FUNCTION_BLOCK UCT_PreTratamento (* UCT Fast de tratamento preliminar + bomba de gordura - HidrycoLib *)
  (* Standard: 61499-2 *)
  (* Version 1.8, 12/11/2026, Hidryco, Hidryco, 1.8: termica da BombaGordura de volta a NF (cfgTermicaNF = TRUE: FALSE no campo = atuada), a pedido do usuario depois de corrigir os nomes dos symlinks (Pre_Tratamento1/2). 1.7: termica da BombaGordura invertida a pedido do usuario (cfgTermicaNF = FALSE: TRUE no campo = atuada). 1.6: IThis.STS_LIGADO, STS_AUTOMATICO (IO List da Nereda). 1.5: eventos da peneira rotativa na logica certa (liga manual em REQ_PEN_LIGA, velocidade em REQ_PEN_VEL, intermitente em REQ_PEN_INT). 1.4: simbolo sGordura (tanque de gordura e valvula de lavagem) para a tela do pre-tratamento. 1.3: sSkid reorganizado (tubos atras, equipamentos alinhados as portas), SymbolSize nos simbolos. 1.2: simbolo sSkid (desenho ISA-101 do skid, com os simbolos dos equipamentos e da bomba de gordura). 1.0: UCT Fast (tratamento preliminar, memorial PR-809) por Modbus TCP. Leitura pela configuracao de hardware (MODBUSGENTCPS + MODBUSRREG8/2 em 40005, 40013, 40081, 40101, 40116, 40127, 40136, 40151, 40161, 40230, 40500, 40508, 40516) nos symlinks ${PATH}mbW005..mbH517 (INT) e connStatusInt em ${PATH}mbConexao; escrita por MODBUSWREG1 em requestwrite nos symlinks ${PATH}mbEscW005..mbEscW017 e ${PATH}mbEscV101..mbEscV161 (INT), so quando o operador comanda. Equipamentos (sub-CATs UCT_Equipamento): Peneira, Bomba1, Bomba2, Valvula1, Valvula2, Compressor, Raspador, Rosca1, Rosca2. Disponibilidade pelo AND editavel (AND_UCT_OK e AND_DISPONIVEL); cadeia antHabilitada/antDisponivel -> stsBloqueioEEE. Bomba de gordura 200-BR-0x (Motor_Generico BombaGordura: E/S por ${PATH}BombaGordura.stsLocal/... e ATV: ComStatus direto em ${PATH}BombaGordura.stsFalhaComunicacao, o motor inverte) e valvula de lavagem ${PATH}cmdValvulaLavagem (BOOL). *)
  PACKAGE Hidryco.HidrycoLib;
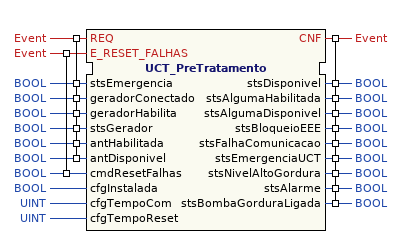
  EVENT_INPUT
    REQ WITH stsEmergencia, geradorConectado, geradorHabilita, stsGerador, antHabilitada, antDisponivel; (* Atualizacao do processo *)
    E_RESET_FALHAS WITH cmdResetFalhas; (* Reset pelo processo (UCT e bomba de gordura) com cmdResetFalhas = TRUE *)
  END_EVENT
  EVENT_OUTPUT
    CNF WITH stsDisponivel, stsAlgumaHabilitada, stsAlgumaDisponivel, stsBloqueioEEE, stsFalhaComunicacao, stsEmergenciaUCT, stsNivelAltoGordura, stsAlarme, stsBombaGorduraLigada; (* Disponibilidade, cadeia das UCTs e estados (so na mudanca) *)
  END_EVENT
  VAR_INPUT
    stsEmergencia : BOOL; (* Emergencia pelo processo: retira o comando da bomba de gordura e fecha a valvula de lavagem *)
    geradorConectado : BOOL := TRUE; (* A bomba de gordura pode ser alimentada pelo gerador *)
    geradorHabilita : BOOL; (* Bomba de gordura liberada para operar com a planta no gerador (HAB_UCT_200_0x do CAT Subestacao) *)
    stsGerador : BOOL; (* Planta alimentada pelo gerador *)
    antHabilitada : BOOL; (* Cadeia: alguma UCT anterior habilitada (stsAlgumaHabilitada da UCT anterior) *)
    antDisponivel : BOOL; (* Cadeia: alguma UCT anterior disponivel (stsAlgumaDisponivel da UCT anterior) *)
    cmdResetFalhas : BOOL; (* TRUE = reset (com o evento E_RESET_FALHAS) *)
    cfgInstalada : BOOL := TRUE; (* FALSE = UCT ainda nao existe em campo (sem comunicacao, sem alarmes, fora do bloqueio da EEE) *)
    cfgTempoCom : UINT := 10; (* Tempo (s) sem comunicacao com a UCT para confirmar a falha *)
    cfgTempoReset : UINT := 2; (* Tempo (s) do pulso de reset escrito na UCT (40005.3) *)
  END_VAR
  VAR_OUTPUT
    stsDisponivel : BOOL; (* UCT disponivel (saida do AND) *)
    stsAlgumaHabilitada : BOOL; (* Esta UCT ou alguma anterior habilitada *)
    stsAlgumaDisponivel : BOOL; (* Esta UCT ou alguma anterior disponivel *)
    stsBloqueioEEE : BOOL; (* Bloqueio do automatico da EEE Bruto: ha UCT habilitada e nenhuma disponivel *)
    stsFalhaComunicacao : BOOL; (* Falha de comunicacao com a UCT *)
    stsEmergenciaUCT : BOOL; (* Emergencia acionada na UCT *)
    stsNivelAltoGordura : BOOL; (* Nivel alto do tanque de gordura (UCT) *)
    stsAlarme : BOOL; (* Algum alarme da UCT *)
    stsBombaGorduraLigada : BOOL; (* Bomba de gordura ligada *)
  END_VAR
  FBS
    IThis : UCT_PreTratamento_HMI(QI := TRUE);
    plcStart1 : plcStart(Prio := 10);
    Logica : basicUCT;
    Tick : E_CYCLE(DT := T#1s);
    Leitura1 : SYMLINKMULTIVARDST_115C998103CD7017B(NAME1 := '$${PATH}mbW005', NAME2 := '$${PATH}mbW006', NAME3 := '$${PATH}mbW007', NAME4 := '$${PATH}mbW008', NAME5 := '$${PATH}mbW009', NAME6 := '$${PATH}mbW010', NAME7 := '$${PATH}mbW011', NAME8 := '$${PATH}mbW012', NAME9 := '$${PATH}mbW013', NAME10 := '$${PATH}mbW014', NAME11 := '$${PATH}mbW015', NAME12 := '$${PATH}mbW016', NAME13 := '$${PATH}mbW017', NAME14 := '$${PATH}mbW081', NAME15 := '$${PATH}mbW082', QI := TRUE); {SET_ATTRIBUTE(Configuration.GenericFBType.InterfaceParams, Runtime.System#I:=15;VALUE${I$}:INT,INT,INT,INT,INT,INT,INT,INT,INT,INT,INT,INT,INT,INT,INT)}
    Leitura2 : SYMLINKMULTIVARDST_115C998103CD7017B(NAME1 := '$${PATH}mbS101', NAME2 := '$${PATH}mbS106', NAME3 := '$${PATH}mbS116', NAME4 := '$${PATH}mbS117', NAME5 := '$${PATH}mbS121', NAME6 := '$${PATH}mbS122', NAME7 := '$${PATH}mbS127', NAME8 := '$${PATH}mbS132', NAME9 := '$${PATH}mbS136', NAME10 := '$${PATH}mbS137', NAME11 := '$${PATH}mbS141', NAME12 := '$${PATH}mbS142', NAME13 := '$${PATH}mbS151', NAME14 := '$${PATH}mbS152', NAME15 := '$${PATH}mbS161', QI := TRUE); {SET_ATTRIBUTE(Configuration.GenericFBType.InterfaceParams, Runtime.System#I:=15;VALUE${I$}:INT,INT,INT,INT,INT,INT,INT,INT,INT,INT,INT,INT,INT,INT,INT)}
    Leitura3 : SYMLINKMULTIVARDST_115C998103CD7017B(NAME1 := '$${PATH}mbS162', NAME2 := '$${PATH}mbW230', NAME3 := '$${PATH}mbH500', NAME4 := '$${PATH}mbH501', NAME5 := '$${PATH}mbH502', NAME6 := '$${PATH}mbH503', NAME7 := '$${PATH}mbH504', NAME8 := '$${PATH}mbH505', NAME9 := '$${PATH}mbH506', NAME10 := '$${PATH}mbH507', NAME11 := '$${PATH}mbH508', NAME12 := '$${PATH}mbH509', NAME13 := '$${PATH}mbH510', NAME14 := '$${PATH}mbH511', NAME15 := '$${PATH}mbH512', QI := TRUE); {SET_ATTRIBUTE(Configuration.GenericFBType.InterfaceParams, Runtime.System#I:=15;VALUE${I$}:INT,INT,INT,INT,INT,INT,INT,INT,INT,INT,INT,INT,INT,INT,INT)}
    Leitura4 : SYMLINKMULTIVARDST_15292F208F22048C1(NAME1 := '$${PATH}mbH513', NAME2 := '$${PATH}mbH514', NAME3 := '$${PATH}mbH515', NAME4 := '$${PATH}mbH516', QI := TRUE); {SET_ATTRIBUTE(Configuration.GenericFBType.InterfaceParams, Runtime.System#I:=4;VALUE${I$}:INT,INT,INT,INT)}
    Leitura5 : SYMLINKMULTIVARDST_5A03F112CD5D470(NAME1 := '$${PATH}mbH517', QI := TRUE); {SET_ATTRIBUTE(Configuration.GenericFBType.InterfaceParams, Runtime.System#I:=1;VALUE${I$}:INT)}
    Comunicacao : SYMLINKMULTIVARDST_5A03F112CD5D470(NAME1 := '$${PATH}mbConexao', QI := TRUE); {SET_ATTRIBUTE(Configuration.GenericFBType.InterfaceParams, Runtime.System#I:=1;VALUE${I$}:INT)}
    EscreveW005 : SYMLINKMULTIVARSRC_5A03F112CD5D470(NAME1 := '$${PATH}mbEscW005', QI := TRUE); {SET_ATTRIBUTE(Configuration.GenericFBType.InterfaceParams, Runtime.System#I:=1;VALUE${I$}:INT)}
    EscreveW006 : SYMLINKMULTIVARSRC_5A03F112CD5D470(NAME1 := '$${PATH}mbEscW006', QI := TRUE); {SET_ATTRIBUTE(Configuration.GenericFBType.InterfaceParams, Runtime.System#I:=1;VALUE${I$}:INT)}
    EscreveW007 : SYMLINKMULTIVARSRC_5A03F112CD5D470(NAME1 := '$${PATH}mbEscW007', QI := TRUE); {SET_ATTRIBUTE(Configuration.GenericFBType.InterfaceParams, Runtime.System#I:=1;VALUE${I$}:INT)}
    EscreveW008 : SYMLINKMULTIVARSRC_5A03F112CD5D470(NAME1 := '$${PATH}mbEscW008', QI := TRUE); {SET_ATTRIBUTE(Configuration.GenericFBType.InterfaceParams, Runtime.System#I:=1;VALUE${I$}:INT)}
    EscreveW009 : SYMLINKMULTIVARSRC_5A03F112CD5D470(NAME1 := '$${PATH}mbEscW009', QI := TRUE); {SET_ATTRIBUTE(Configuration.GenericFBType.InterfaceParams, Runtime.System#I:=1;VALUE${I$}:INT)}
    EscreveW010 : SYMLINKMULTIVARSRC_5A03F112CD5D470(NAME1 := '$${PATH}mbEscW010', QI := TRUE); {SET_ATTRIBUTE(Configuration.GenericFBType.InterfaceParams, Runtime.System#I:=1;VALUE${I$}:INT)}
    EscreveW011 : SYMLINKMULTIVARSRC_5A03F112CD5D470(NAME1 := '$${PATH}mbEscW011', QI := TRUE); {SET_ATTRIBUTE(Configuration.GenericFBType.InterfaceParams, Runtime.System#I:=1;VALUE${I$}:INT)}
    EscreveW012 : SYMLINKMULTIVARSRC_5A03F112CD5D470(NAME1 := '$${PATH}mbEscW012', QI := TRUE); {SET_ATTRIBUTE(Configuration.GenericFBType.InterfaceParams, Runtime.System#I:=1;VALUE${I$}:INT)}
    EscreveW013 : SYMLINKMULTIVARSRC_5A03F112CD5D470(NAME1 := '$${PATH}mbEscW013', QI := TRUE); {SET_ATTRIBUTE(Configuration.GenericFBType.InterfaceParams, Runtime.System#I:=1;VALUE${I$}:INT)}
    EscreveW014 : SYMLINKMULTIVARSRC_5A03F112CD5D470(NAME1 := '$${PATH}mbEscW014', QI := TRUE); {SET_ATTRIBUTE(Configuration.GenericFBType.InterfaceParams, Runtime.System#I:=1;VALUE${I$}:INT)}
    EscreveW015 : SYMLINKMULTIVARSRC_5A03F112CD5D470(NAME1 := '$${PATH}mbEscW015', QI := TRUE); {SET_ATTRIBUTE(Configuration.GenericFBType.InterfaceParams, Runtime.System#I:=1;VALUE${I$}:INT)}
    EscreveW016 : SYMLINKMULTIVARSRC_5A03F112CD5D470(NAME1 := '$${PATH}mbEscW016', QI := TRUE); {SET_ATTRIBUTE(Configuration.GenericFBType.InterfaceParams, Runtime.System#I:=1;VALUE${I$}:INT)}
    EscreveW017 : SYMLINKMULTIVARSRC_5A03F112CD5D470(NAME1 := '$${PATH}mbEscW017', QI := TRUE); {SET_ATTRIBUTE(Configuration.GenericFBType.InterfaceParams, Runtime.System#I:=1;VALUE${I$}:INT)}
    EscreveV101 : SYMLINKMULTIVARSRC_5A03F112CD5D470(NAME1 := '$${PATH}mbEscV101', QI := TRUE); {SET_ATTRIBUTE(Configuration.GenericFBType.InterfaceParams, Runtime.System#I:=1;VALUE${I$}:INT)}
    EscreveV116 : SYMLINKMULTIVARSRC_5A03F112CD5D470(NAME1 := '$${PATH}mbEscV116', QI := TRUE); {SET_ATTRIBUTE(Configuration.GenericFBType.InterfaceParams, Runtime.System#I:=1;VALUE${I$}:INT)}
    EscreveV121 : SYMLINKMULTIVARSRC_5A03F112CD5D470(NAME1 := '$${PATH}mbEscV121', QI := TRUE); {SET_ATTRIBUTE(Configuration.GenericFBType.InterfaceParams, Runtime.System#I:=1;VALUE${I$}:INT)}
    EscreveV136 : SYMLINKMULTIVARSRC_5A03F112CD5D470(NAME1 := '$${PATH}mbEscV136', QI := TRUE); {SET_ATTRIBUTE(Configuration.GenericFBType.InterfaceParams, Runtime.System#I:=1;VALUE${I$}:INT)}
    EscreveV141 : SYMLINKMULTIVARSRC_5A03F112CD5D470(NAME1 := '$${PATH}mbEscV141', QI := TRUE); {SET_ATTRIBUTE(Configuration.GenericFBType.InterfaceParams, Runtime.System#I:=1;VALUE${I$}:INT)}
    EscreveV151 : SYMLINKMULTIVARSRC_5A03F112CD5D470(NAME1 := '$${PATH}mbEscV151', QI := TRUE); {SET_ATTRIBUTE(Configuration.GenericFBType.InterfaceParams, Runtime.System#I:=1;VALUE${I$}:INT)}
    EscreveV161 : SYMLINKMULTIVARSRC_5A03F112CD5D470(NAME1 := '$${PATH}mbEscV161', QI := TRUE); {SET_ATTRIBUTE(Configuration.GenericFBType.InterfaceParams, Runtime.System#I:=1;VALUE${I$}:INT)}
    ValvulaLavagem : SYMLINKMULTIVARSRC_1559B0FF8170C9BA0(NAME1 := '$${PATH}cmdValvulaLavagem', QI := TRUE); {SET_ATTRIBUTE(Configuration.GenericFBType.InterfaceParams, Runtime.System#I:=1;VALUE${I$}:BOOL)}
    AND_UCT_OK : AND_1122770BAB85676D3; {SET_ATTRIBUTE(Configuration.GenericFBType.InterfaceParams, Runtime.Standard#CNT:=3)}
    AND_DISPONIVEL : AND_1122770BAB85676D3; {SET_ATTRIBUTE(Configuration.GenericFBType.InterfaceParams, Runtime.Standard#CNT:=3)}
    Bomba_Higienizacao1 : UCT_Equipamento(pin_6729E072E11CC02E := TRUE, pin_B3CA2188BE2BF3D0 := FALSE, pin_E5B528FA2A3E5A83 := FALSE);
    Bomba_Higienizacao2 : UCT_Equipamento(pin_6729E072E11CC02E := TRUE, pin_B3CA2188BE2BF3D0 := FALSE, pin_E5B528FA2A3E5A83 := FALSE);
    Valvula_Higienizacao1 : UCT_Equipamento(pin_6729E072E11CC02E := FALSE, pin_B3CA2188BE2BF3D0 := FALSE, pin_E5B528FA2A3E5A83 := FALSE);
    Valvula_Higienizacao2 : UCT_Equipamento(pin_6729E072E11CC02E := FALSE, pin_B3CA2188BE2BF3D0 := FALSE, pin_E5B528FA2A3E5A83 := FALSE);
    Compressor1 : UCT_Equipamento(pin_6729E072E11CC02E := TRUE, pin_B3CA2188BE2BF3D0 := FALSE, pin_E5B528FA2A3E5A83 := FALSE);
    Raspador_Gordura1 : UCT_Equipamento(pin_6729E072E11CC02E := TRUE, pin_B3CA2188BE2BF3D0 := TRUE, pin_E5B528FA2A3E5A83 := TRUE);
    Rosca1Horizontal : UCT_Equipamento(pin_6729E072E11CC02E := TRUE, pin_B3CA2188BE2BF3D0 := TRUE, pin_E5B528FA2A3E5A83 := TRUE);
    Rosca2Inclinada : UCT_Equipamento(pin_6729E072E11CC02E := TRUE, pin_B3CA2188BE2BF3D0 := TRUE, pin_E5B528FA2A3E5A83 := TRUE);
    BombaGordura : Motor_Generico(pin_63EFEFB7C85EC93E := TRUE, pin_66763E13F70A4420 := TRUE, pin_D34C88BE7FFF3208 := TRUE, pin_39489193B7758574 := 600.0);
    AlarmeCom : ALARM_BIT(TYPE := 1, ACKTYPE_1 := 2, ACTIVE := TRUE); {SET_ATTRIBUTE(HMI.AlarmText, UCT sem comunicação)}
    AlarmeEmergencia : ALARM_BIT(TYPE := 1, ACKTYPE_1 := 2, ACTIVE := TRUE); {SET_ATTRIBUTE(HMI.AlarmText, Emergência acionada na UCT)}
    AlarmeDefPEN : ALARM_BIT(TYPE := 1, ACKTYPE_1 := 2, ACTIVE := TRUE); {SET_ATTRIBUTE(HMI.AlarmText, Defeito na peneira rotativa)}
    AlarmeDefB1 : ALARM_BIT(TYPE := 1, ACKTYPE_1 := 2, ACTIVE := TRUE); {SET_ATTRIBUTE(HMI.AlarmText, Defeito na bomba 1 de higienização da peneira)}
    AlarmeDefB2 : ALARM_BIT(TYPE := 1, ACKTYPE_1 := 2, ACTIVE := TRUE); {SET_ATTRIBUTE(HMI.AlarmText, Defeito na bomba 2 de higienização da peneira)}
    AlarmeDefCMP : ALARM_BIT(TYPE := 1, ACKTYPE_1 := 2, ACTIVE := TRUE); {SET_ATTRIBUTE(HMI.AlarmText, Defeito no compressor de ar)}
    AlarmeDefRSP : ALARM_BIT(TYPE := 1, ACKTYPE_1 := 2, ACTIVE := TRUE); {SET_ATTRIBUTE(HMI.AlarmText, Defeito no raspador de gordura)}
    AlarmeDefR1 : ALARM_BIT(TYPE := 1, ACKTYPE_1 := 2, ACTIVE := TRUE); {SET_ATTRIBUTE(HMI.AlarmText, Defeito na rosca 1 (horizontal))}
    AlarmeDefR2 : ALARM_BIT(TYPE := 1, ACKTYPE_1 := 2, ACTIVE := TRUE); {SET_ATTRIBUTE(HMI.AlarmText, Defeito na rosca 2 (inclinada))}
    AlarmeNivelAgua : ALARM_BIT(TYPE := 1, ACKTYPE_1 := 2, ACTIVE := TRUE); {SET_ATTRIBUTE(HMI.AlarmText, Nível baixo no tanque de água de higienização)} {SET_ATTRIBUTE(HMI.AlarmClass, Warning)}
    AlarmeNivelPeneira : ALARM_BIT(TYPE := 1, ACKTYPE_1 := 2, ACTIVE := TRUE); {SET_ATTRIBUTE(HMI.AlarmText, Nível alto na peneira)} {SET_ATTRIBUTE(HMI.AlarmClass, Warning)}
    Peneira_Rotativa1 : UCT_Equipamento(pin_6729E072E11CC02E := TRUE, pin_B3CA2188BE2BF3D0 := TRUE, pin_E5B528FA2A3E5A83 := FALSE);
  END_FBS
  EVENT_CONNECTIONS
    plcStart1.FIRST_INIT TO IThis.7731B1FFA94C6332;
    plcStart1.REDO_INIT TO IThis.7731B1FFA94C6332;
    IThis.BE90C28BEC8DBAC0 TO Logica.3C5B6DD981EA9EF0;
    Logica.416B84A41F220B84 TO Tick.START;
    Logica.416B84A41F220B84 TO Leitura1.INIT;
    Logica.416B84A41F220B84 TO Leitura2.INIT;
    Logica.416B84A41F220B84 TO Leitura3.INIT;
    Logica.416B84A41F220B84 TO Leitura4.INIT;
    Logica.416B84A41F220B84 TO Leitura5.INIT;
    Logica.416B84A41F220B84 TO Comunicacao.INIT;
    Logica.416B84A41F220B84 TO EscreveW005.INIT;
    Logica.416B84A41F220B84 TO EscreveW006.INIT;
    Logica.416B84A41F220B84 TO EscreveW007.INIT;
    Logica.416B84A41F220B84 TO EscreveW008.INIT;
    Logica.416B84A41F220B84 TO EscreveW009.INIT;
    Logica.416B84A41F220B84 TO EscreveW010.INIT;
    Logica.416B84A41F220B84 TO EscreveW011.INIT;
    Logica.416B84A41F220B84 TO EscreveW012.INIT;
    Logica.416B84A41F220B84 TO EscreveW013.INIT;
    Logica.416B84A41F220B84 TO EscreveW014.INIT;
    Logica.416B84A41F220B84 TO EscreveW015.INIT;
    Logica.416B84A41F220B84 TO EscreveW016.INIT;
    Logica.416B84A41F220B84 TO EscreveW017.INIT;
    Logica.416B84A41F220B84 TO EscreveV101.INIT;
    Logica.416B84A41F220B84 TO EscreveV116.INIT;
    Logica.416B84A41F220B84 TO EscreveV121.INIT;
    Logica.416B84A41F220B84 TO EscreveV136.INIT;
    Logica.416B84A41F220B84 TO EscreveV141.INIT;
    Logica.416B84A41F220B84 TO EscreveV151.INIT;
    Logica.416B84A41F220B84 TO EscreveV161.INIT;
    Logica.416B84A41F220B84 TO ValvulaLavagem.INIT;
    Logica.416B84A41F220B84 TO AlarmeCom.INIT;
    AlarmeCom.INITO TO AlarmeCom.REQ_INITDATA;
    AlarmeCom.CNF_INITDATA TO AlarmeCom.ACTIVATE;
    AlarmeCom.INITO TO AlarmeEmergencia.INIT;
    AlarmeEmergencia.INITO TO AlarmeEmergencia.REQ_INITDATA;
    AlarmeEmergencia.CNF_INITDATA TO AlarmeEmergencia.ACTIVATE;
    AlarmeEmergencia.INITO TO AlarmeDefPEN.INIT;
    AlarmeDefPEN.INITO TO AlarmeDefPEN.REQ_INITDATA;
    AlarmeDefPEN.CNF_INITDATA TO AlarmeDefPEN.ACTIVATE;
    AlarmeDefPEN.INITO TO AlarmeDefB1.INIT;
    AlarmeDefB1.INITO TO AlarmeDefB1.REQ_INITDATA;
    AlarmeDefB1.CNF_INITDATA TO AlarmeDefB1.ACTIVATE;
    AlarmeDefB1.INITO TO AlarmeDefB2.INIT;
    AlarmeDefB2.INITO TO AlarmeDefB2.REQ_INITDATA;
    AlarmeDefB2.CNF_INITDATA TO AlarmeDefB2.ACTIVATE;
    AlarmeDefB2.INITO TO AlarmeDefCMP.INIT;
    AlarmeDefCMP.INITO TO AlarmeDefCMP.REQ_INITDATA;
    AlarmeDefCMP.CNF_INITDATA TO AlarmeDefCMP.ACTIVATE;
    AlarmeDefCMP.INITO TO AlarmeDefRSP.INIT;
    AlarmeDefRSP.INITO TO AlarmeDefRSP.REQ_INITDATA;
    AlarmeDefRSP.CNF_INITDATA TO AlarmeDefRSP.ACTIVATE;
    AlarmeDefRSP.INITO TO AlarmeDefR1.INIT;
    AlarmeDefR1.INITO TO AlarmeDefR1.REQ_INITDATA;
    AlarmeDefR1.CNF_INITDATA TO AlarmeDefR1.ACTIVATE;
    AlarmeDefR1.INITO TO AlarmeDefR2.INIT;
    AlarmeDefR2.INITO TO AlarmeDefR2.REQ_INITDATA;
    AlarmeDefR2.CNF_INITDATA TO AlarmeDefR2.ACTIVATE;
    AlarmeDefR2.INITO TO AlarmeNivelAgua.INIT;
    AlarmeNivelAgua.INITO TO AlarmeNivelAgua.REQ_INITDATA;
    AlarmeNivelAgua.CNF_INITDATA TO AlarmeNivelAgua.ACTIVATE;
    AlarmeNivelAgua.INITO TO AlarmeNivelPeneira.INIT;
    AlarmeNivelPeneira.INITO TO AlarmeNivelPeneira.REQ_INITDATA;
    AlarmeNivelPeneira.CNF_INITDATA TO AlarmeNivelPeneira.ACTIVATE;
    AlarmeNivelPeneira.INITO TO plcStart1.ACK_FIRST;
    AlarmeNivelPeneira.INITO TO IThis.BF3BAA6EB0D69F6F;
    Leitura1.CNF TO Logica.86B21E575F925410;
    Leitura2.CNF TO Logica.ACF117E29FC3AC1C;
    Leitura3.CNF TO Logica.FD034B0BBE440D40;
    Leitura4.CNF TO Logica.729388FCDFDF68AE;
    Leitura5.CNF TO Logica.96AC3F0A2629C81D;
    Comunicacao.CNF TO Logica.4327DB3EB2D5D05C;
    Logica.11F41745985917DF TO EscreveW005.REQ;
    Logica.E9DD31896C582136 TO EscreveW006.REQ;
    Logica.E928AC62D8378E2E TO EscreveW007.REQ;
    Logica.8C6CC9C5F833000C TO EscreveW008.REQ;
    Logica.10A819F294BECD61 TO EscreveW009.REQ;
    Logica.CCE6CEE36384A6FD TO EscreveW010.REQ;
    Logica.48F5F46EFA41CB2E TO EscreveW011.REQ;
    Logica.FB2D821A4BBF6B61 TO EscreveW012.REQ;
    Logica.6F9E0D27072C9DCA TO EscreveW013.REQ;
    Logica.3830C851999B1CA8 TO EscreveW014.REQ;
    Logica.91DFFB362B8ECB72 TO EscreveW015.REQ;
    Logica.D8E5B77061056FA5 TO EscreveW016.REQ;
    Logica.67B496F21A680217 TO EscreveW017.REQ;
    Logica.2DC67FC3F907B62C TO EscreveV101.REQ;
    Logica.9697531BFDFDAA11 TO EscreveV116.REQ;
    Logica.EA10A30027EF1458 TO EscreveV121.REQ;
    Logica.76B63473D5644862 TO EscreveV136.REQ;
    Logica.E8A88BE3B83ED632 TO EscreveV141.REQ;
    Logica.FCC1975F18BB837D TO EscreveV151.REQ;
    Logica.D44CECCDCDAFDF05 TO EscreveV161.REQ;
    Logica.8621D711C765D74F TO ValvulaLavagem.REQ;
    Logica.A0C13DD0452107CB TO Bomba_Higienizacao1.70A516C5CA4155CA;
    Bomba_Higienizacao1.0ECDAB45E7B0C5AF TO Logica.9D9E81ADADCAA296;
    Bomba_Higienizacao1.2D7A148B2A7AA879 TO Logica.E34661574BF84379;
    Logica.A0C13DD0452107CB TO Bomba_Higienizacao2.70A516C5CA4155CA;
    Bomba_Higienizacao2.0ECDAB45E7B0C5AF TO Logica.D87E7B2D8E293BB6;
    Bomba_Higienizacao2.2D7A148B2A7AA879 TO Logica.7CA1C2A34CD31341;
    Logica.A0C13DD0452107CB TO Valvula_Higienizacao1.70A516C5CA4155CA;
    Valvula_Higienizacao1.0ECDAB45E7B0C5AF TO Logica.CF56824B76A4E51B;
    Logica.A0C13DD0452107CB TO Valvula_Higienizacao2.70A516C5CA4155CA;
    Valvula_Higienizacao2.0ECDAB45E7B0C5AF TO Logica.F75EA032D1A6B02C;
    Logica.A0C13DD0452107CB TO Compressor1.70A516C5CA4155CA;
    Compressor1.0ECDAB45E7B0C5AF TO Logica.548C5ECAC6439F23;
    Compressor1.2D7A148B2A7AA879 TO Logica.D33EB6DFF7EADA48;
    Logica.A0C13DD0452107CB TO Raspador_Gordura1.70A516C5CA4155CA;
    Raspador_Gordura1.0ECDAB45E7B0C5AF TO Logica.4F24C39CA1B377DA;
    Raspador_Gordura1.453EBF0958E76CD5 TO Logica.25A416A6D88DD0BD;
    Raspador_Gordura1.D9A88CBEE21DBA8E TO Logica.2DDC9EB582C567B6;
    Raspador_Gordura1.2D7A148B2A7AA879 TO Logica.E445565C572BE9AB;
    Logica.A0C13DD0452107CB TO Rosca1Horizontal.70A516C5CA4155CA;
    Rosca1Horizontal.0ECDAB45E7B0C5AF TO Logica.B6026660A2849366;
    Rosca1Horizontal.453EBF0958E76CD5 TO Logica.38389BFD6E07A057;
    Rosca1Horizontal.D9A88CBEE21DBA8E TO Logica.460B0CE006F8F781;
    Rosca1Horizontal.2D7A148B2A7AA879 TO Logica.9798AA2801C41B49;
    Logica.A0C13DD0452107CB TO Rosca2Inclinada.70A516C5CA4155CA;
    Rosca2Inclinada.0ECDAB45E7B0C5AF TO Logica.05FCFC0A4F34DAC5;
    Rosca2Inclinada.453EBF0958E76CD5 TO Logica.917F967EEA65C256;
    Rosca2Inclinada.D9A88CBEE21DBA8E TO Logica.F6429B88CEB00ADB;
    Rosca2Inclinada.2D7A148B2A7AA879 TO Logica.66FC9636E69253EA;
    IThis.1F1F8302525DDF94 TO Logica.60A9FA7D1B9019D9;
    IThis.1EA45A01E944042C TO Logica.10C669586AF9B729;
    IThis.6BDBFED6495F25F4 TO Logica.70D47E2D73B66C31;
    IThis.734C7A77C68CFD95 TO Logica.10434994C0931297;
    IThis.E2F5EBA7E91047EB TO Logica.4287AE5C00B681B1;
    IThis.CA131EB7F5B48041 TO Logica.8858219971D3BAD6;
    IThis.09F2CE520A7CB40A TO Logica.B055BD39F7E10E53;
    IThis.74FD7728297A1739 TO Logica.8B3CC5BA21742708;
    IThis.36C4ED263F60138F TO Logica.01DDB779929E0BD3;
    IThis.313AA7AFD2DEA98C TO Logica.FF42D335F0EB104F;
    E_RESET_FALHAS TO Logica.F6EC819575FB3804;
    REQ TO Logica.75410FBD6637F3BE;
    REQ TO BombaGordura.21070E4B73BFECDC;
    Tick.EO TO Logica.41222487C8D9CF7D;
    Logica.A4E8AA815C7798D0 TO CNF;
    Logica.B1173782F7B0D885 TO IThis.4D2C1FBBFC38ACE6;
    Logica.4C6FF34A6B3F84FA TO AND_UCT_OK.REQ;
    AND_UCT_OK.CNF TO AND_DISPONIVEL.REQ;
    AND_DISPONIVEL.CNF TO Logica.B4B1263914B085C1;
    Logica.31FE10FED34E3AE0 TO BombaGordura.21070E4B73BFECDC;
    BombaGordura.9D4F26EE27EDF5B9 TO Logica.7F4121B3EAF345EF;
    BombaGordura.9D4F26EE27EDF5B9 TO CNF;
    Logica.61B5851DEAB87FC2 TO BombaGordura.BA30A65ADDA4ECC3;
    Logica.B2C6B3F912408F66 TO AlarmeCom.REQ;
    Logica.B2C6B3F912408F66 TO AlarmeEmergencia.REQ;
    Logica.B2C6B3F912408F66 TO AlarmeDefPEN.REQ;
    Logica.B2C6B3F912408F66 TO AlarmeDefB1.REQ;
    Logica.B2C6B3F912408F66 TO AlarmeDefB2.REQ;
    Logica.B2C6B3F912408F66 TO AlarmeDefCMP.REQ;
    Logica.B2C6B3F912408F66 TO AlarmeDefRSP.REQ;
    Logica.B2C6B3F912408F66 TO AlarmeDefR1.REQ;
    Logica.B2C6B3F912408F66 TO AlarmeDefR2.REQ;
    Logica.B2C6B3F912408F66 TO AlarmeNivelAgua.REQ;
    Logica.B2C6B3F912408F66 TO AlarmeNivelPeneira.REQ;
    AlarmeCom.IND_1 TO IThis.4D2C1FBBFC38ACE6;
    AlarmeEmergencia.IND_1 TO IThis.4D2C1FBBFC38ACE6;
    AlarmeDefPEN.IND_1 TO IThis.4D2C1FBBFC38ACE6;
    AlarmeDefB1.IND_1 TO IThis.4D2C1FBBFC38ACE6;
    AlarmeDefB2.IND_1 TO IThis.4D2C1FBBFC38ACE6;
    AlarmeDefCMP.IND_1 TO IThis.4D2C1FBBFC38ACE6;
    AlarmeDefRSP.IND_1 TO IThis.4D2C1FBBFC38ACE6;
    AlarmeDefR1.IND_1 TO IThis.4D2C1FBBFC38ACE6;
    AlarmeDefR2.IND_1 TO IThis.4D2C1FBBFC38ACE6;
    AlarmeNivelAgua.IND_1 TO IThis.4D2C1FBBFC38ACE6;
    AlarmeNivelPeneira.IND_1 TO IThis.4D2C1FBBFC38ACE6;
    IThis.74FD7728297A1739 TO AlarmeCom.ACK_C1;
    IThis.74FD7728297A1739 TO AlarmeEmergencia.ACK_C1;
    IThis.74FD7728297A1739 TO AlarmeDefPEN.ACK_C1;
    IThis.74FD7728297A1739 TO AlarmeDefB1.ACK_C1;
    IThis.74FD7728297A1739 TO AlarmeDefB2.ACK_C1;
    IThis.74FD7728297A1739 TO AlarmeDefCMP.ACK_C1;
    IThis.74FD7728297A1739 TO AlarmeDefRSP.ACK_C1;
    IThis.74FD7728297A1739 TO AlarmeDefR1.ACK_C1;
    IThis.74FD7728297A1739 TO AlarmeDefR2.ACK_C1;
    IThis.74FD7728297A1739 TO AlarmeNivelAgua.ACK_C1;
    IThis.74FD7728297A1739 TO AlarmeNivelPeneira.ACK_C1;
    E_RESET_FALHAS TO AlarmeCom.ACK_C1;
    E_RESET_FALHAS TO AlarmeEmergencia.ACK_C1;
    E_RESET_FALHAS TO AlarmeDefPEN.ACK_C1;
    E_RESET_FALHAS TO AlarmeDefB1.ACK_C1;
    E_RESET_FALHAS TO AlarmeDefB2.ACK_C1;
    E_RESET_FALHAS TO AlarmeDefCMP.ACK_C1;
    E_RESET_FALHAS TO AlarmeDefRSP.ACK_C1;
    E_RESET_FALHAS TO AlarmeDefR1.ACK_C1;
    E_RESET_FALHAS TO AlarmeDefR2.ACK_C1;
    E_RESET_FALHAS TO AlarmeNivelAgua.ACK_C1;
    E_RESET_FALHAS TO AlarmeNivelPeneira.ACK_C1;
    Logica.A4E8AA815C7798D0 TO Peneira_Rotativa1.70A516C5CA4155CA;
    Logica.B1173782F7B0D885 TO Peneira_Rotativa1.70A516C5CA4155CA;
    Logica.A0C13DD0452107CB TO Peneira_Rotativa1.70A516C5CA4155CA;
    Logica.4C6FF34A6B3F84FA TO Peneira_Rotativa1.70A516C5CA4155CA;
    Logica.B2C6B3F912408F66 TO Peneira_Rotativa1.70A516C5CA4155CA;
    Logica.31FE10FED34E3AE0 TO Peneira_Rotativa1.70A516C5CA4155CA;
    Logica.8621D711C765D74F TO Peneira_Rotativa1.70A516C5CA4155CA;
    Logica.61B5851DEAB87FC2 TO Peneira_Rotativa1.70A516C5CA4155CA;
    Peneira_Rotativa1.0ECDAB45E7B0C5AF TO Logica.F5A0AE6E537529F5;
    Peneira_Rotativa1.2D7A148B2A7AA879 TO Logica.4A489282C873CE35;
    Peneira_Rotativa1.453EBF0958E76CD5 TO Logica.CB1FF06E5DD10F71;
  END_CONNECTIONS
  DATA_CONNECTIONS
    cfgInstalada TO Logica.B84AF20A00A0FEAB;
    cfgTempoCom TO Logica.2D0DECC616DD4E29;
    cfgTempoReset TO Logica.6F72EF7A9957D9B1;
    cmdResetFalhas TO Logica.F64D45B3992C3082;
    antHabilitada TO Logica.CF63D4AF765659C1;
    antDisponivel TO Logica.9756EA9EC3EE5693;
    stsEmergencia TO Logica.BCC8272ACE7AC349;
    Leitura1.VALUE1 TO Logica.2AF241D1E0537909;
    Leitura1.VALUE2 TO Logica.EB87F4844550BF0A;
    Leitura1.VALUE3 TO Logica.702CACE592B586EC;
    Leitura1.VALUE4 TO Logica.00E434C4D2FCE1E2;
    Leitura1.VALUE5 TO Logica.216DC8D1B0130B70;
    Leitura1.VALUE6 TO Logica.E92E8124C98345A8;
    Leitura1.VALUE7 TO Logica.5702FCE80FD9232F;
    Leitura1.VALUE8 TO Logica.2C198397DC93FDE4;
    Leitura1.VALUE9 TO Logica.8DC0D656670A81AF;
    Leitura1.VALUE10 TO Logica.FF2A6CB505BDEEED;
    Leitura1.VALUE11 TO Logica.29D39A9131350120;
    Leitura1.VALUE12 TO Logica.5047554D33D25508;
    Leitura1.VALUE13 TO Logica.6213901E687BF582;
    Leitura1.VALUE14 TO Logica.805F5AA59EEEC2D4;
    Leitura1.VALUE15 TO Logica.8AF7D7600739FBD8;
    Leitura2.VALUE1 TO Logica.CBA17D927032CBD4;
    Leitura2.VALUE2 TO Logica.E81009FF89B5BC15;
    Leitura2.VALUE3 TO Logica.FDB62ADC45542E9E;
    Leitura2.VALUE4 TO Logica.6D9544B2D05EE83A;
    Leitura2.VALUE5 TO Logica.EAC2F7A409142C5D;
    Leitura2.VALUE6 TO Logica.2873DE3B6BFE44C9;
    Leitura2.VALUE7 TO Logica.DB13AC717A8B7662;
    Leitura2.VALUE8 TO Logica.4D5D876EB3A7F171;
    Leitura2.VALUE9 TO Logica.51DA211617F1996B;
    Leitura2.VALUE10 TO Logica.97151C90B367E8DC;
    Leitura2.VALUE11 TO Logica.EEFE5F1EF8383B49;
    Leitura2.VALUE12 TO Logica.62F04539174C591F;
    Leitura2.VALUE13 TO Logica.02097632451711DE;
    Leitura2.VALUE14 TO Logica.7991843F9B2D5590;
    Leitura2.VALUE15 TO Logica.DDA25525CB8A7B4D;
    Leitura3.VALUE1 TO Logica.111326FFB7350BF0;
    Leitura3.VALUE2 TO Logica.605236348EF76178;
    Leitura3.VALUE3 TO Logica.009C88AD569306A2;
    Leitura3.VALUE4 TO Logica.A0B989F0831D5C46;
    Leitura3.VALUE5 TO Logica.C7387B9A6FCCB81F;
    Leitura3.VALUE6 TO Logica.E47649B3DC153190;
    Leitura3.VALUE7 TO Logica.3553691F126CE1B5;
    Leitura3.VALUE8 TO Logica.0A36A58BDBBC0471;
    Leitura3.VALUE9 TO Logica.42520E00029B280F;
    Leitura3.VALUE10 TO Logica.B3A245D474F32D30;
    Leitura3.VALUE11 TO Logica.FDF3C709AEBF1C84;
    Leitura3.VALUE12 TO Logica.25EE4A659CDB8B19;
    Leitura3.VALUE13 TO Logica.8E1D474EDFE3E373;
    Leitura3.VALUE14 TO Logica.A05F827665BFFF1E;
    Leitura3.VALUE15 TO Logica.DE0C347B4E1AA668;
    Leitura4.VALUE1 TO Logica.BE7F6B173ECEF46F;
    Leitura4.VALUE2 TO Logica.5FDC3C3D54E86285;
    Leitura4.VALUE3 TO Logica.D1FE5B095A8ACDE9;
    Leitura4.VALUE4 TO Logica.8A95E69557A2E9BE;
    Leitura5.VALUE1 TO Logica.ED8792C392F4F103;
    Comunicacao.VALUE1 TO Logica.8E65120B34D38BDE;
    Logica.48B51513B83DEAC1 TO EscreveW005.VALUE1;
    Logica.ABE25A7B6D246024 TO EscreveW006.VALUE1;
    Logica.332BB6C4B414C757 TO EscreveW007.VALUE1;
    Logica.5FF35C3FF4051574 TO EscreveW008.VALUE1;
    Logica.7BCA7ABE5B2A80CB TO EscreveW009.VALUE1;
    Logica.EE8A41D2485DFDB4 TO EscreveW010.VALUE1;
    Logica.A2EA9BE38D7D6BAA TO EscreveW011.VALUE1;
    Logica.126C934AB0F6DBFE TO EscreveW012.VALUE1;
    Logica.73DD8991441412AC TO EscreveW013.VALUE1;
    Logica.DE2C0333DCDCC77C TO EscreveW014.VALUE1;
    Logica.8B46394DF76CFFD8 TO EscreveW015.VALUE1;
    Logica.B5B936F289F2140E TO EscreveW016.VALUE1;
    Logica.96F874CA969849BC TO EscreveW017.VALUE1;
    Logica.93EC120EF49D8A9B TO EscreveV101.VALUE1;
    Logica.B84F5A34C7CB0F43 TO EscreveV116.VALUE1;
    Logica.2EEB0ECC5C70DFC8 TO EscreveV121.VALUE1;
    Logica.A95766D7DCAD36EA TO EscreveV136.VALUE1;
    Logica.D451279D5E50FC08 TO EscreveV141.VALUE1;
    Logica.D04BD37BABA3A53F TO EscreveV151.VALUE1;
    Logica.77B5D89A59E485CC TO EscreveV161.VALUE1;
    Logica.97A930D5B8996F70 TO ValvulaLavagem.VALUE1;
    Logica.4FE6015A2477CFC9 TO AND_UCT_OK.IN1;
    Logica.3836FD4FBDBFBB63 TO AND_UCT_OK.IN2;
    Logica.CFDFC80ABF4D39D0 TO AND_UCT_OK.IN3;
    AND_UCT_OK.OUT TO AND_DISPONIVEL.IN1;
    Logica.9719C72C2028949E TO AND_DISPONIVEL.IN2;
    Logica.EAECF18552174CCF TO AND_DISPONIVEL.IN3;
    AND_DISPONIVEL.OUT TO Logica.907F6462227B081B;
    Logica.9F5A0BAAA6BA36FB TO Bomba_Higienizacao1.93B31B867A532500;
    Logica.B0882E75048E56C8 TO Bomba_Higienizacao1.98FD5EAA90BD9629;
    Logica.F433D77752764E72 TO Bomba_Higienizacao1.96E48787F8AC58C3;
    Logica.BB50EA5A17772016 TO Bomba_Higienizacao1.CC220F735371196B;
    Logica.6D499885ADD13F89 TO Bomba_Higienizacao1.33285C93B9AAB2BC;
    Logica.6F1E502C9B6CF2B2 TO Bomba_Higienizacao1.3F39B194DE4581AB;
    Logica.B8856E3515E1335F TO Bomba_Higienizacao1.F6AE4997ED76CC8B;
    Logica.48FD745C0144715F TO Bomba_Higienizacao1.0E2695E0A2003068;
    Bomba_Higienizacao1.074D328E856330C0 TO Logica.C19AEC3805E7291E;
    Bomba_Higienizacao1.520AB5A4EADBD8AE TO Logica.878937D8CA59CE95;
    Logica.26DA29A2F44AB1D9 TO Bomba_Higienizacao2.93B31B867A532500;
    Logica.AE4A01B00246A9BC TO Bomba_Higienizacao2.98FD5EAA90BD9629;
    Logica.49B62932E0024FCB TO Bomba_Higienizacao2.96E48787F8AC58C3;
    Logica.C62B70166A0883C7 TO Bomba_Higienizacao2.CC220F735371196B;
    Logica.3229D99A95CB4D5D TO Bomba_Higienizacao2.33285C93B9AAB2BC;
    Logica.AC94358F5B25F765 TO Bomba_Higienizacao2.3F39B194DE4581AB;
    Logica.8F6F2CB2BBCF9FC3 TO Bomba_Higienizacao2.F6AE4997ED76CC8B;
    Logica.4FF14F19D4AA0DEA TO Bomba_Higienizacao2.0E2695E0A2003068;
    Bomba_Higienizacao2.074D328E856330C0 TO Logica.6F688A786E95C4D1;
    Bomba_Higienizacao2.520AB5A4EADBD8AE TO Logica.3A9274E19001885E;
    Logica.9594942602D571EA TO Valvula_Higienizacao1.93B31B867A532500;
    Logica.3A38DC7CA6958C9C TO Valvula_Higienizacao1.98FD5EAA90BD9629;
    Logica.3E823B19B09A5097 TO Valvula_Higienizacao1.96E48787F8AC58C3;
    Logica.13E9E7335A7C2901 TO Valvula_Higienizacao1.CC220F735371196B;
    Logica.A66FC5515667CF08 TO Valvula_Higienizacao1.33285C93B9AAB2BC;
    Logica.3FD3C8118B86508A TO Valvula_Higienizacao1.3F39B194DE4581AB;
    Logica.ACC893CA1C181DB0 TO Valvula_Higienizacao1.F6AE4997ED76CC8B;
    Logica.3B6C8D4012CD67E8 TO Valvula_Higienizacao1.0E2695E0A2003068;
    Valvula_Higienizacao1.074D328E856330C0 TO Logica.E44BA349DE6CBE3D;
    Logica.83D44C4C3C2A69C6 TO Valvula_Higienizacao2.93B31B867A532500;
    Logica.2ADE61FFCD947701 TO Valvula_Higienizacao2.98FD5EAA90BD9629;
    Logica.AB418D0D39BCD6F9 TO Valvula_Higienizacao2.96E48787F8AC58C3;
    Logica.214258657E323579 TO Valvula_Higienizacao2.CC220F735371196B;
    Logica.2205641E77B9A34C TO Valvula_Higienizacao2.33285C93B9AAB2BC;
    Logica.B8A2E15DD4914861 TO Valvula_Higienizacao2.3F39B194DE4581AB;
    Logica.608E639AB4ED2F8D TO Valvula_Higienizacao2.F6AE4997ED76CC8B;
    Logica.7DAD37347BA7821F TO Valvula_Higienizacao2.0E2695E0A2003068;
    Valvula_Higienizacao2.074D328E856330C0 TO Logica.90EFC5FA870ED8B5;
    Logica.4B03E2982EF25D75 TO Compressor1.93B31B867A532500;
    Logica.9A133A3818AB7D75 TO Compressor1.98FD5EAA90BD9629;
    Logica.894358E3DD02DC60 TO Compressor1.96E48787F8AC58C3;
    Logica.04D5D6C179AAB7E5 TO Compressor1.CC220F735371196B;
    Logica.684C8B722280E4D3 TO Compressor1.33285C93B9AAB2BC;
    Logica.C315013255DF205C TO Compressor1.3F39B194DE4581AB;
    Logica.5ECE4DBB763DBD73 TO Compressor1.F6AE4997ED76CC8B;
    Logica.5C65E619BE12DEDB TO Compressor1.0E2695E0A2003068;
    Compressor1.074D328E856330C0 TO Logica.3ECA38388FA33BAB;
    Compressor1.520AB5A4EADBD8AE TO Logica.54782A528428A27E;
    Logica.8C265EEC37B1503A TO Raspador_Gordura1.93B31B867A532500;
    Logica.10B9DDCA13A25793 TO Raspador_Gordura1.98FD5EAA90BD9629;
    Logica.7D6D39D384DEE9A7 TO Raspador_Gordura1.96E48787F8AC58C3;
    Logica.2665663CA7E8C4E3 TO Raspador_Gordura1.CC220F735371196B;
    Logica.ECB4D30DAD3A8F7A TO Raspador_Gordura1.33285C93B9AAB2BC;
    Logica.80173FD5AD234274 TO Raspador_Gordura1.3F39B194DE4581AB;
    Logica.67FEABF9507CF440 TO Raspador_Gordura1.F6AE4997ED76CC8B;
    Logica.CFD27D979F18C5A5 TO Raspador_Gordura1.0E2695E0A2003068;
    Raspador_Gordura1.074D328E856330C0 TO Logica.EF5E268AEC8FFB6F;
    Raspador_Gordura1.C49C9947FE6383D2 TO Logica.CD033E2BD625D117;
    Raspador_Gordura1.E18D01D6E7CD5F0A TO Logica.ABC0CD4591666DED;
    Raspador_Gordura1.520AB5A4EADBD8AE TO Logica.C50C1B75AA3833A4;
    Logica.A972128A35D56662 TO Rosca1Horizontal.93B31B867A532500;
    Logica.62F4E28E677AF90C TO Rosca1Horizontal.98FD5EAA90BD9629;
    Logica.F84A9EFD3BC7F02B TO Rosca1Horizontal.96E48787F8AC58C3;
    Logica.7307C4B442730619 TO Rosca1Horizontal.CC220F735371196B;
    Logica.B624A1A3392B6721 TO Rosca1Horizontal.33285C93B9AAB2BC;
    Logica.EC246D0019464C9A TO Rosca1Horizontal.3F39B194DE4581AB;
    Logica.8530A93EC6E0B63B TO Rosca1Horizontal.F6AE4997ED76CC8B;
    Logica.970B608B8836000A TO Rosca1Horizontal.0E2695E0A2003068;
    Rosca1Horizontal.074D328E856330C0 TO Logica.3BCA796FB5DBD06E;
    Rosca1Horizontal.C49C9947FE6383D2 TO Logica.F95CCCF398D56F2E;
    Rosca1Horizontal.E18D01D6E7CD5F0A TO Logica.2227D73D7FD55805;
    Rosca1Horizontal.520AB5A4EADBD8AE TO Logica.5CEF29EA4AD62820;
    Logica.08E4196F96764545 TO Rosca2Inclinada.93B31B867A532500;
    Logica.2EBC40C7F99057D2 TO Rosca2Inclinada.98FD5EAA90BD9629;
    Logica.A91E1AB8D5A774D8 TO Rosca2Inclinada.96E48787F8AC58C3;
    Logica.EFC6255887164B86 TO Rosca2Inclinada.CC220F735371196B;
    Logica.0268E3B1CAFAE678 TO Rosca2Inclinada.33285C93B9AAB2BC;
    Logica.F0652198FBD98A9C TO Rosca2Inclinada.3F39B194DE4581AB;
    Logica.531FF78EC4DA12AC TO Rosca2Inclinada.F6AE4997ED76CC8B;
    Logica.25E9EBFC2025D937 TO Rosca2Inclinada.0E2695E0A2003068;
    Rosca2Inclinada.074D328E856330C0 TO Logica.2C67200E4B5EFF53;
    Rosca2Inclinada.C49C9947FE6383D2 TO Logica.411B151F745A6FE5;
    Rosca2Inclinada.E18D01D6E7CD5F0A TO Logica.F7464DBF7DB7632E;
    Rosca2Inclinada.520AB5A4EADBD8AE TO Logica.C9BA77924D8D8C4A;
    IThis.E8EC0002033C76CE TO Logica.679AB85673B231F7;
    IThis.6D865A5A332E5543 TO Logica.597C737D269B71D2;
    IThis.BF399167056A87ED TO Logica.174D0C5CEEEE344F;
    IThis.77BCED6C06D331DF TO Logica.C4A8663B0D52BA34;
    IThis.17E93345B45473CC TO Logica.C21FD557DB2DAA26;
    IThis.F2302575AAD84B02 TO Logica.6BFC54B0FFB9A684;
    IThis.4EFF59B0E8A8A572 TO Logica.B940523A960C2800;
    IThis.57D3892FB897956D TO Logica.07B2B2CF770F4814;
    IThis.E01817B0B9D294F0 TO Logica.E8439982309E033C;
    IThis.BC3F99BD918D681D TO Logica.D48C361677C598B3;
    IThis.7E14DCADCFEAB7FC TO Logica.9BC9AEB7EE8B0E7A;
    IThis.74687B9042CE2260 TO Logica.969BCD5D8972BBD3;
    IThis.9D4C68BE8DF350DA TO Logica.48C7D048A8BBA01A;
    IThis.557377A1B5F4A834 TO Logica.4471CCC90EDB124D;
    Logica.3FCEA38A9E6EE5CE TO BombaGordura.87DAE15414E7C412;
    Logica.370D92A80C450D03 TO BombaGordura.F94ABA993E8E9FF4;
    stsEmergencia TO BombaGordura.85953C7B9294A9BF;
    geradorConectado TO BombaGordura.8914049066EE23D9;
    geradorHabilita TO BombaGordura.5C3D51A654AD25BA;
    stsGerador TO BombaGordura.A33BC24B3E7310B0;
    Logica.EB86EA91F4C64D64 TO BombaGordura.C2F1E9C0FB076F17;
    BombaGordura.40A5976BFB296133 TO Logica.E35B723AAFA80B5D;
    BombaGordura.368C3F9EC04E0359 TO Logica.13F60FFCABA8441A;
    BombaGordura.40A5976BFB296133 TO stsBombaGorduraLigada;
    Logica.7F7B816331BE1C2B TO AlarmeCom.INP;
    Logica.3614F51665280D43 TO AlarmeEmergencia.INP;
    Logica.145A4BA522A4B16C TO AlarmeDefPEN.INP;
    Logica.350AC8442CDE22A1 TO AlarmeDefB1.INP;
    Logica.AFE2F9492D389BBD TO AlarmeDefB2.INP;
    Logica.798FABD1834C18CD TO AlarmeDefCMP.INP;
    Logica.CAD3C184BA624DED TO AlarmeDefRSP.INP;
    Logica.8C0378D10BE98D49 TO AlarmeDefR1.INP;
    Logica.78B77585A68CAB67 TO AlarmeDefR2.INP;
    Logica.C76BC1CB5B2AF8A0 TO AlarmeNivelAgua.INP;
    Logica.FD8522ED9B351538 TO AlarmeNivelPeneira.INP;
    Logica.578D8BBF4DA79A23 TO stsDisponivel;
    Logica.84171C035357B4E3 TO stsAlgumaHabilitada;
    Logica.B1E45CD679DEB114 TO stsAlgumaDisponivel;
    Logica.D73E486392D4D5B6 TO stsBloqueioEEE;
    Logica.C0D9728386F92C77 TO stsFalhaComunicacao;
    Logica.EB99489D8453BA21 TO stsEmergenciaUCT;
    Logica.37ECE09B1E5AEFFB TO stsNivelAltoGordura;
    Logica.FA37E7894F6BD3D0 TO stsAlarme;
    Logica.EB99489D8453BA21 TO IThis.77996B129DEED446;
    Logica.0647910676F94640 TO IThis.C66C21CCD4DB83C0;
    Logica.F3713950EE5D1867 TO IThis.337E31D7EDB8F44A;
    Logica.7D2A38C25D8FD93C TO IThis.9C9347BCFEAF7AF9;
    Logica.37ECE09B1E5AEFFB TO IThis.E4136C8F6C1D00EC;
    Logica.C4EE1E8A3DAA5B83 TO IThis.2952D3783A30100B;
    Logica.C0D9728386F92C77 TO IThis.424CD593158BAD0D;
    Logica.578D8BBF4DA79A23 TO IThis.7FC922186689F6A7;
    Logica.EAECF18552174CCF TO IThis.F2EEAD9F89C10C0A;
    Logica.D73E486392D4D5B6 TO IThis.DB03AD759AC99D87;
    Logica.FA37E7894F6BD3D0 TO IThis.0754132ADEC84B47;
    Logica.642EE6D10F9115A0 TO IThis.8DB404409CDC4860;
    Logica.B8C76428B99C0BC3 TO IThis.1E5F0BD6663A26A0;
    Logica.4C8B357E982AEFA5 TO IThis.34CA8296753C9B57;
    Logica.42BCE54FED382E40 TO IThis.FD3EE3853B4F44E7;
    Logica.3C697FA38E7B1CEE TO IThis.5C6534C9699DB5B6;
    Logica.35B9945971456169 TO IThis.A34EAF033F42F954;
    Logica.DDCDDDAAC0A5E903 TO IThis.5313A39E74F246C2;
    Logica.D1AFC6808E3F4248 TO IThis.53C171BAA75F8591;
    Logica.98BD502D5E024892 TO IThis.7DD1B5310A9624B5;
    Logica.74B9486C9619CFB9 TO IThis.12C80A903AD4A502;
    Logica.7F7B816331BE1C2B TO IThis.656FE051A422C54F;
    Logica.3614F51665280D43 TO IThis.6712AE6DDCBDA2C3;
    Logica.145A4BA522A4B16C TO IThis.FE92207488FBF5FB;
    Logica.350AC8442CDE22A1 TO IThis.EC56E017B9BDB5F3;
    Logica.AFE2F9492D389BBD TO IThis.4A9DF66D259412E5;
    Logica.798FABD1834C18CD TO IThis.1F68FD40C57BEF36;
    Logica.CAD3C184BA624DED TO IThis.396053A9E11344C5;
    Logica.8C0378D10BE98D49 TO IThis.F107E2325FA54130;
    Logica.78B77585A68CAB67 TO IThis.BF05A8169FEC3401;
    Logica.C76BC1CB5B2AF8A0 TO IThis.8FD364E4C6F826F0;
    Logica.FD8522ED9B351538 TO IThis.E5B8FA1CAB955B70;
    AlarmeCom.STATE_1 TO IThis.236E5D50753D714E;
    AlarmeEmergencia.STATE_1 TO IThis.5F1046313EDB69DC;
    AlarmeDefPEN.STATE_1 TO IThis.7A71B775DFFE9B1C;
    AlarmeDefB1.STATE_1 TO IThis.0E08B20C4ED421EB;
    AlarmeDefB2.STATE_1 TO IThis.48AC31BF354006CB;
    AlarmeDefCMP.STATE_1 TO IThis.DE8D247CD85A57E5;
    AlarmeDefRSP.STATE_1 TO IThis.B1CD278E523A9C55;
    AlarmeDefR1.STATE_1 TO IThis.084992A935E4A85E;
    AlarmeDefR2.STATE_1 TO IThis.CDD01305047A1ACC;
    AlarmeNivelAgua.STATE_1 TO IThis.A8C53509FE285DA7;
    AlarmeNivelPeneira.STATE_1 TO IThis.1D197D0EC16DF374;
    Logica.E15602DD5EFD812C TO Peneira_Rotativa1.93B31B867A532500;
    Logica.895BD8D8326C37F1 TO Peneira_Rotativa1.98FD5EAA90BD9629;
    Logica.71216940FF3AAA09 TO Peneira_Rotativa1.96E48787F8AC58C3;
    Logica.431ACF2EB10AEC5B TO Peneira_Rotativa1.CC220F735371196B;
    Logica.FCE2010BC99734E0 TO Peneira_Rotativa1.33285C93B9AAB2BC;
    Logica.82C23DAE5245FE05 TO Peneira_Rotativa1.3F39B194DE4581AB;
    Logica.4EAFAAC987F7E6ED TO Peneira_Rotativa1.F6AE4997ED76CC8B;
    Logica.630B3326E520DED3 TO Peneira_Rotativa1.0E2695E0A2003068;
    Peneira_Rotativa1.074D328E856330C0 TO Logica.19CB07B401748599;
    Peneira_Rotativa1.520AB5A4EADBD8AE TO Logica.368D14EA4B585390;
    Peneira_Rotativa1.C49C9947FE6383D2 TO Logica.4EB5BC958EA12D54;
    Logica.65044E21F1507E93 TO IThis.19EF5D97B246D865;
    Logica.642EE6D10F9115A0 TO IThis.911C06B9DECB84C5;
  END_CONNECTIONS
END_FUNCTION_BLOCK
